Fanuc KAREL source: kt00883.KL

-- PROVISIONAL review KL for V770-1; original PC SHA256 61cecebbcf3dbef8a5650b03c208319c7629e8e208cd45e79a34077898f7c96a
-- Incomplete behavior may be omitted. Consult companion uncertainty JSON. Do not deploy.
PROGRAM KT00883
%NOLOCKGROUP
VAR
  R1 : REAL
  R2 : REAL
  OUT : REAL
BEGIN
  -- UNRESOLVED_PC offsets 5-16; opcodes 2E,23
  -- UNRESOLVED_PC offsets 21-32; opcodes 2E,23
  -- UNRESOLVED_PC offsets 37-48; opcodes 2E,23
  -- UNRESOLVED_PC offsets 53-64; opcodes 2E,23
  -- UNRESOLVED_PC offsets 69-90; opcodes 27,22,22,76,23
  -- UNRESOLVED_PC offsets 95-99; opcodes 7F
END KT00883
